                num nSigType[3]
                num nValue[3]
            mdesc mMdesc = {leave=0}
            num nActionIndex = 60
            num nDelay = 1
            num nMoveType = 1
            num nPercentage
            num nSigValue = 1
        pointRx pPointRx[2] = {x=-138.850367, y=-44.569058, z=962.511805, rx=-1.752214, ry=-0.122124, rz=-89.326646, shoulder=lefty, elbow=epositive, wrist=wpositive}
        string sID
      [75]
        bool bMarked
        jointRx jJointRx = {j1=-49.904251, j2=-65.605747, j3=139.0621971, j4=-181.0710428, j5=74.878861, j6=140.871685}
        pointRx pInter
        paraItem pParaItem
          [0]
            bool bSafePoint
            ifItem iIfItem
              [0]
                bool bANDOR[2]
                num nSigIndex[3]
                num nSigType[3]
                num nValue[3]
            mdesc mMdesc = {leave=0}
            num nActionIndex = 60
            num nDelay = 1
            num nMoveType = 1
            num nPercentage
            num nSigValue = 1
        pointRx pPointRx[2] = {x=-44.539892, y=-44.568217, z=962.547058, rx=-1.752061, ry=-0.123361, rz=-89.326689, shoulder=lefty, elbow=epositive, wrist=wpositive}
        string sID
      [76]
        bool bMarked
        jointRx jJointRx = {j1=-49.289261, j2=-63.229169, j3=134.202102, j4=-181.102758, j5=72.384398, j6=140.311025}
        pointRx pInter
        paraItem pParaItem
          [0]
            bool bSafePoint
            ifItem iIfItem
              [0]
                bool bANDOR[2]
                num nSigIndex[3]
                num nSigType[3]
                num nValue[3]
            mdesc mMdesc = {leave=0}
            num nActionIndex = 60
            num nDelay = 1
            num nMoveType = 1
            num nPercentage
            num nSigValue = 1
        pointRx pPointRx[2] = {x=-42.782853, y=-44.569273, z=1003.955298, rx=-1.753071, ry=-0.121713, rz=-89.326781, shoulder=lefty, elbow=epositive, wrist=wpositive}
        string sID
      [77]
        bool bMarked
        jointRx jJointRx = {j1=-25.432487, j2=-45.494499, j3=127.259364, j4=-181.493414, j5=82.715062, j6=116.303511}
        pointRx pInter
        paraItem pParaItem
          [0]
            bool bSafePoint
            ifItem iIfItem
              [0]
                bool bANDOR[2]
                num nSigIndex[3]
                num nSigType[3]
                num nValue[3]
            mdesc mMdesc = {leave=0}
            num nActionIndex = 60
            num nDelay = 1
            num nMoveType = 1
            num nPercentage
            num nSigValue = 1
        pointRx pPointRx[2] = {x=73.884399, y=-40.550183, z=1028.430042, rx=-1.744787, ry=-0.219486, rz=-89.333983, shoulder=lefty, elbow=epositive, wrist=wpositive}
        string sID
      [78]
        bool bMarked
        jointRx jJointRx = {j1=-57.856377, j2=-66.18455, j3=133.138862, j4=-180.798841, j5=68.549304, j6=148.828951}
        pointRx pInter
        paraItem pParaItem
          [0]
            bool bSafePoint
            ifItem iIfItem
              [0]
                bool bANDOR[2]
                num nSigIndex[3]
                num nSigType[3]
                num nValue[3]
            mdesc mMdesc = {leave=0}
            num nActionIndex = 60
            num nDelay = 1
            num nMoveType = 1
            num nPercentage
            num nSigValue = 1
        pointRx pPointRx[2] = {x=-67.43152, y=-40.567065, z=1016.367875, rx=-1.744462, ry=-0.217896, rz=-89.333233, shoulder=lefty, elbow=epositive, wrist=wpositive}
        string sID
      [79]
        bool bMarked
        jointRx jJointRx = {j1=-125.666138, j2=-76.447258, j3=135.218346, j4=-178.621352, j5=60.0693288, j6=215.6343}
        pointRx pInter
        paraItem pParaItem
          [0]
            bool bSafePoint
            ifItem iIfItem
              [0]
                bool bANDOR[2]
                num nSigIndex[3]
                num nSigType[3]
                num nValue[3]
            mdesc mMdesc = {leave=0}
            num nActionIndex = 60
            num nDelay = 1
            num nMoveType = 1
            num nPercentage
            num nSigValue = 1
        pointRx pPointRx[2] = {x=-141.607559, y=-40.56496, z=1001.487797, rx=-1.745427, ry=-0.218033, rz=-89.333718, shoulder=lefty, elbow=epositive, wrist=wpositive}
        string sID
      [80]
        bool bMarked
        jointRx jJointRx = {j1=-163.468753, j2=-72.941717, j3=129.657925, j4=-177.930129, j5=57.0209808, j6=253.00669774}
        pointRx pInter
        paraItem pParaItem
          [0]
            bool bSafePoint
            ifItem iIfItem
              [0]
                bool bANDOR[2]
                num nSigIndex[3]
                num nSigType[3]
                num nValue[3]
            mdesc mMdesc = {leave=0}
            num nActionIndex = 60
            num nDelay = 1
            num nMoveType = 1
            num nPercentage
            num nSigValue = 1
        pointRx pPointRx[2] = {x=-178.509464, y=-40.567787, z=1047.669101, rx=-1.746323, ry=-0.218277, rz=-89.333981, shoulder=lefty, elbow=epositive, wrist=wpositive}
        string sID
      [81]
        bool bMarked
        jointRx jJointRx = {j1=-177.244487, j2=-58.712757, j3=130.795458, j4=-178.155232, j5=71.95685, j6=267.344536}
        pointRx pInter
        paraItem pParaItem
          [0]
            bool bSafePoint
            ifItem iIfItem
              [0]
                bool bANDOR[2]
                num nSigIndex[3]
                num nSigType[3]
                num nValue[3]
            mdesc mMdesc = {leave=0}
            num nActionIndex = 60
            num nDelay = 1
            num nMoveType = 1
            num nPercentage
            num nSigValue = 1
        pointRx pPointRx[2] = {x=-305.74421, y=-40.564807, z=1028.0320815, rx=-1.745533, ry=-0.218693, rz=-89.333779, shoulder=lefty, elbow=epositive, wrist=wpositive}
        string sID
      [82]
        bool bMarked
        jointRx jJointRx = {j1=-178.526843, j2=-40.454962, j3=125.405301, j4=-178.242312, j5=84.778901, j6=269.0391142}
        pointRx pInter
        paraItem pParaItem
          [0]
            bool bSafePoint
            ifItem iIfItem
              [0]
                bool bANDOR[2]
                num nSigIndex[3]
                num nSigType[3]
                num nValue[3]
            mdesc mMdesc = {leave=0}
            num nActionIndex = 60
            num nDelay = 1
            num nMoveType = 1
            num nPercentage
            num nSigValue = 1
        pointRx pPointRx[2] = {x=-434.343088, y=-40.61718, z=1028.0320848, rx=-1.745356, ry=-0.218738, rz=-89.333719, shoulder=lefty, elbow=epositive, wrist=wpositive}
        string sID
      [83]
        bool bMarked
        jointRx jJointRx = {j1=-178.966416, j2=-24.85944, j3=117.444048, j4=-178.24946, j5=92.396091, j6=269.712104}
        pointRx pInter
        paraItem pParaItem
          [0]
            bool bSafePoint
            ifItem iIfItem
              [0]
                bool bANDOR[2]
                num nSigIndex[3]
                num nSigType[3]
                num nValue[3]
            mdesc mMdesc = {leave=0}
            num nActionIndex = 60
            num nDelay = 1
            num nMoveType = 1
            num nPercentage
            num nSigValue = 1
        pointRx pPointRx[2] = {x=-550.558, y=-40.617172, z=1028.0320539, rx=-1.745357, ry=-0.218827, rz=-89.333714, shoulder=lefty, elbow=epositive, wrist=wpositive}
        string sID
      [84]
        bool bMarked
        jointRx jJointRx = {j1=-178.990337, j2=-23.604156, j3=109.459463, j4=-178.246238, j5=85.670511, j6=269.530325}
        pointRx pInter
        paraItem pParaItem
          [0]
            bool bSafePoint
            ifItem iIfItem
              [0]
                bool bANDOR[2]
                num nSigIndex[3]
                num nSigType[3]
                num nValue[3]
            mdesc mMdesc = {leave=0}
            num nActionIndex = 60
            num nDelay = 1
            num nMoveType = 1
            num nPercentage
            num nSigValue = 1
        pointRx pPointRx[2] = {x=-559.676751, y=-40.616999, z=1097.0852879, rx=-1.745205, ry=-0.217512, rz=-89.33374, shoulder=lefty, elbow=epositive, wrist=wpositive}
        string sID
      [85]
        bool bMarked
        jointRx jJointRx = {j1=-178.943744, j2=-24.322013, j3=101.711175, j4=-178.206641, j5=77.210582, j6=269.219034}
        pointRx pInter
        paraItem pParaItem
          [0]
            bool bSafePoint
            ifItem iIfItem
              [0]
                bool bANDOR[2]
                num nSigIndex[3]
                num nSigType[3]
                num nValue[3]
            mdesc mMdesc = {leave=0}
            num nActionIndex = 60
            num nDelay = 1
            num nMoveType = 1
            num nPercentage
            num nSigValue = 1
        pointRx pPointRx[2] = {x=-542.070783, y=-40.616994, z=1174.87195, rx=-1.745164, ry=-0.216758, rz=-89.333713, shoulder=lefty, elbow=epositive, wrist=wpositive}
        string sID
      [86]
        bool bMarked
        jointRx jJointRx = {j1=-178.943806, j2=-23.793943, j3=99.30263, j4=-178.192287, j5=75.331347, j6=269.158327}
        pointRx pInter
        paraItem pParaItem
          [0]
            bool bSafePoint
            ifItem iIfItem
              [0]
                bool bANDOR[2]
                num nSigIndex[3]
                num nSigType[3]
                num nValue[3]
            mdesc mMdesc = {leave=0}
            num nActionIndex = 60
            num nDelay = 1
            num nMoveType = 1
            num nPercentage
            num nSigValue = 1
        pointRx pPointRx[2] = {x=-542.046055, y=-40.616997, z=1194.299438, rx=-1.745092, ry=-0.216442, rz=-89.333682, shoulder=lefty, elbow=epositive, wrist=wpositive}
        string sID
      [87]
        bool bMarked
        jointRx jJointRx = {j1=-178.85922, j2=-27.330123, j3=102.744036, j4=-178.191054, j5=75.238753, j6=269.0705123}
        pointRx pInter
        paraItem pParaItem
          [0]
            bool bSafePoint
            ifItem iIfItem
              [0]
                bool bANDOR[2]
                num nSigIndex[3]
                num nSigType[3]
                num nValue[3]
            mdesc mMdesc = {leave=0}
            num nActionIndex = 60
            num nDelay = 1
            num nMoveType = 1
            num nPercentage
            num nSigValue = 1
        pointRx pPointRx[2] = {x=-513.909364, y=-40.617001, z=1181.865557, rx=-1.745263, ry=-0.216897, rz=-89.333745, shoulder=lefty, elbow=epositive, wrist=wpositive}
        string sID
      [88]
        bool bMarked
        jointRx jJointRx = {j1=-178.577868, j2=-35.0352996, j3=106.0927297, j4=-178.147828, j5=70.89347, j6=268.643627}
        pointRx pInter
        paraItem pParaItem
          [0]
            bool bSafePoint
            ifItem iIfItem
              [0]
                bool bANDOR[2]
                num nSigIndex[3]
                num nSigType[3]
                num nValue[3]
            mdesc mMdesc = {leave=0}
            num nActionIndex = 60
            num nDelay = 1
            num nMoveType = 1
            num nPercentage
            num nSigValue = 1
        pointRx pPointRx[2] = {x=-444.101189, y=-40.617001, z=1187.110134, rx=-1.745281, ry=-0.216517, rz=-89.333733, shoulder=lefty, elbow=epositive, wrist=wpositive}
        string sID
      [89]
        bool bMarked
        jointRx jJointRx = {j1=-177.964362, j2=-47.427804, j3=117.345153, j4=-178.132839, j5=69.773165, j6=267.990525}
        pointRx pInter
        paraItem pParaItem
          [0]
            bool bSafePoint
            ifItem iIfItem
              [0]
                bool bANDOR[2]
                num nSigIndex[3]
                num nSigType[3]
                num nValue[3]
            mdesc mMdesc = {leave=0}
            num nActionIndex = 60
            num nDelay = 1
            num nMoveType = 1
            num nPercentage
            num nSigValue = 1
        pointRx pPointRx[2] = {x=-358.696243, y=-40.617001, z=1126.286618, rx=-1.745413, ry=-0.216112, rz=-89.333736, shoulder=lefty, elbow=epositive, wrist=wpositive}
        string sID
      [90]
        bool bMarked
        jointRx jJointRx = {j1=-177.960401, j2=-42.42338, j3=104.324192, j4=-178.0116171, j5=61.761954, j6=267.691309}
        pointRx pInter
        paraItem pParaItem
          [0]
            bool bSafePoint
            ifItem iIfItem
              [0]
                bool bANDOR[2]
                num nSigIndex[3]
                num nSigType[3]
                num nValue[3]
            mdesc mMdesc = {leave=0}
            num nActionIndex = 60
            num nDelay = 1
            num nMoveType = 1
            num nPercentage
            num nSigValue = 1
        pointRx pPointRx[2] = {x=-358.210554, y=-40.616999, z=1227.312647, rx=-1.745114, ry=-0.215409, rz=-89.333647, shoulder=lefty, elbow=epositive, wrist=wpositive}
        string sID
      [91]
        bool bMarked
        jointRx jJointRx = {j1=-157.648785, j2=-55.0873266, j3=110.653004, j4=-177.95404, j5=56.0449416, j6=247.169842}
        pointRx pInter
        paraItem pParaItem
          [0]
            bool bSafePoint
            ifItem iIfItem
              [0]
                bool bANDOR[2]
                num nSigIndex[3]
                num nSigType[3]
                num nValue[3]
            mdesc mMdesc = {leave=0}
            num nActionIndex = 60
            num nDelay = 1
            num nMoveType = 1
            num nPercentage
            num nSigValue = 1
        pointRx pPointRx[2] = {x=-229.83526, y=-65.451897, z=1196.333444, rx=-1.745262, ry=-0.217825, rz=-89.332323, shoulder=lefty, elbow=epositive, wrist=wpositive}
        string sID
      [92]
        bool bMarked
        jointRx jJointRx = {j1=-152.966394, j2=-56.240625, j3=110.746536, j4=-177.982817, j5=55.121987, j6=242.474574}
        pointRx pInter
        paraItem pParaItem
          [0]
            bool bSafePoint
            ifItem iIfItem
              [0]
                bool bANDOR[2]
                num nSigIndex[3]
                num nSigType[3]
                num nValue[3]
            mdesc mMdesc = {leave=0}
            num nActionIndex = 60
            num nDelay = 1
            num nMoveType = 1
            num nPercentage
            num nSigValue = 1
        pointRx pPointRx[2] = {x=-212.6845, y=-65.452346, z=1196.358042, rx=-1.746333, ry=-0.218302, rz=-89.332682, shoulder=lefty, elbow=epositive, wrist=wpositive}
        string sID
      [93]
        bool bMarked
        jointRx jJointRx = {j1=-118.542599, j2=-58.519116, j3=112.0638486, j4=-178.749072, j5=54.980609, j6=208.482941}
        pointRx pInter
        paraItem pParaItem
          [0]
            bool bSafePoint
            ifItem iIfItem
              [0]
                bool bANDOR[2]
                num nSigIndex[3]
                num nSigType[3]
                num nValue[3]
            mdesc mMdesc = {leave=0}
            num nActionIndex = 60
            num nDelay = 1
            num nMoveType = 1
            num nPercentage
            num nSigValue = 1
        pointRx pPointRx[2] = {x=-149.858699, y=-65.452346, z=1187.0826994, rx=-1.745135, ry=-0.217044, rz=-89.332258, shoulder=lefty, elbow=epositive, wrist=wpositive}
        string sID
      [94]
        bool bMarked
        jointRx jJointRx = {j1=-101.200662, j2=-58.679642, j3=113.706302, j4=-179.339305, j5=56.697308, j6=191.500759}
        pointRx pInter
        paraItem pParaItem
          [0]
            bool bSafePoint
            ifItem iIfItem
              [0]
                bool bANDOR[2]
                num nSigIndex[3]
                num nSigType[3]
                num nValue[3]
            mdesc mMdesc = {leave=0}
            num nActionIndex = 60
            num nDelay = 1
            num nMoveType = 1
            num nPercentage
            num nSigValue = 1
        pointRx pPointRx[2] = {x=-127.503998, y=-65.472867, z=1174.335896, rx=-1.744346, ry=-0.217552, rz=-89.332398, shoulder=lefty, elbow=epositive, wrist=wpositive}
        string sID
      [95]
        bool bMarked
        jointRx jJointRx = {j1=-101.203749, j2=-57.0328969, j3=110.693044, j4=-179.328951, j5=55.331019, j6=191.484931}
        pointRx pInter
        paraItem pParaItem
          [0]
            bool bSafePoint
            ifItem iIfItem
              [0]
                bool bANDOR[2]
                num nSigIndex[3]
                num nSigType[3]
                num nValue[3]
            mdesc mMdesc = {leave=0}
            num nActionIndex = 60
            num nDelay = 1
            num nMoveType = 1
            num nPercentage
            num nSigValue = 1
        pointRx pPointRx[2] = {x=-127.503988, y=-65.473043, z=1197.162512, rx=-1.744433, ry=-0.217146, rz=-89.332357, shoulder=lefty, elbow=epositive, wrist=wpositive}
        string sID
      [96]
        bool bMarked
        jointRx jJointRx = {j1=-84.916197, j2=-57.654127, j3=112.0354709, j4=-179.926433, j5=56.138092, j6=175.545215}
        pointRx pInter
        paraItem pParaItem
          [0]
            bool bSafePoint
            ifItem iIfItem
              [0]
                bool bANDOR[2]
                num nSigIndex[3]
                num nSigType[3]
                num nValue[3]
            mdesc mMdesc = {leave=0}
            num nActionIndex = 60
            num nDelay = 1
            num nMoveType = 1
            num nPercentage
            num nSigValue = 1
        pointRx pPointRx[2] = {x=-105.833813, y=-53.577317, z=1186.997866, rx=-1.744409, ry=-0.216493, rz=-89.33235, shoulder=lefty, elbow=epositive, wrist=wpositive}
        string sID
      [97]
        bool bMarked
        jointRx jJointRx = {j1=-74.942351, j2=-49.0636516, j3=113.425459, j4=-183.373141, j5=77.590842, j6=166.743204}
        pointRx pInter
        paraItem pParaItem
          [0]
            bool bSafePoint
            ifItem iIfItem
              [0]
                bool bANDOR[2]
                num nSigIndex[3]
                num nSigType[3]
                num nValue[3]
            mdesc mMdesc = {leave=0}
            num nActionIndex = 60
            num nDelay = 1
            num nMoveType = 1
            num nPercentage
            num nSigValue = 1
        pointRx pPointRx[2] = {x=-70.288394, y=-10.197743, z=1148.602795, rx=-13.604008, ry=-0.216042, rz=-89.332075, shoulder=lefty, elbow=epositive, wrist=wpositive}
        string sID
      [98]
        bool bMarked
        jointRx jJointRx = {j1=-22.441628, j2=-49.998667, j3=113.146837, j4=-179.268601, j5=63.114949, j6=112.777772}
        pointRx pInter
        paraItem pParaItem
          [0]
            bool bSafePoint
            ifItem iIfItem
              [0]
                bool bANDOR[2]
                num nSigIndex[3]
                num nSigType[3]
                num nValue[3]
            mdesc mMdesc = {leave=0}
            num nActionIndex = 60
            num nDelay = 1
            num nMoveType = 1
            num nPercentage
            num nSigValue = 1
        pointRx pPointRx[2] = {x=2.572536, y=-22.293277, z=1169.165569, rx=0.616343, ry=-0.216579, rz=-89.332136, shoulder=lefty, elbow=epositive, wrist=wpositive}
        string sID
      [99]
        bool bMarked
        jointRx jJointRx = {j1=-16.222078, j2=-42.747965, j3=111.131068, j4=-179.299489, j5=68.420107, j6=106.63085}
        pointRx pInter
        paraItem pParaItem
          [0]
            bool bSafePoint
            ifItem iIfItem
              [0]
                bool bANDOR[2]
                num nSigIndex[3]
                num nSigType[3]
                num nValue[3]
            mdesc mMdesc = {leave=0}
            num nActionIndex = 60
            num nDelay = 1
            num nMoveType = 1
            num nPercentage
            num nSigValue = 1
        pointRx pPointRx[2] = {x=64.811204, y=-22.293322, z=1169.130311, rx=0.615547, ry=-0.216097, rz=-89.332208, shoulder=lefty, elbow=epositive, wrist=wpositive}
        string sID
      [100]
        bool bMarked
        jointRx jJointRx = {j1=-11.927651, j2=-32.0900118, j3=103.0810682, j4=-179.315894, j5=71.0760377, j6=102.371735}
        pointRx pInter
        paraItem pParaItem
          [0]
            bool bSafePoint
            ifItem iIfItem
              [0]
                bool bANDOR[2]
                num nSigIndex[3]
                num nSigType[3]
                num nValue[3]
            mdesc mMdesc = {leave=0}
            num nActionIndex = 60
            num nDelay = 1
            num nMoveType = 1
            num nPercentage
            num nSigValue = 1
        pointRx pPointRx[2] = {x=145.897455, y=-22.29476, z=1202.0898265, rx=0.615855, ry=-0.215659, rz=-89.332409, shoulder=lefty, elbow=epositive, wrist=wpositive}
        string sID
      [101]
        bool bMarked
        jointRx jJointRx = {j1=-14.974019, j2=-36.733975, j3=99.744873, j4=-179.269184, j5=63.0625851, j6=105.309151}
        pointRx pInter
        paraItem pParaItem
          [0]
            bool bSafePoint
            ifItem iIfItem
              [0]
                bool bANDOR[2]
                num nSigIndex[3]
                num nSigType[3]
                num nValue[3]
            mdesc mMdesc = {leave=0}
            num nActionIndex = 60
            num nDelay = 1
            num nMoveType = 1
            num nPercentage
            num nSigValue = 1
        pointRx pPointRx[2] = {x=83.529929, y=-22.294757, z=1249.648683, rx=0.616531, ry=-0.216447, rz=-89.332334, shoulder=lefty, elbow=epositive, wrist=wpositive}
        string sID
      [102]
        bool bMarked
        jointRx jJointRx = {j1=-14.974848, j2=-34.297369, j3=93.572735, j4=-179.243247, j5=59.326428, j6=105.254901}
        pointRx pInter
        paraItem pParaItem
          [0]
            bool bSafePoint
            ifItem iIfItem
              [0]
                bool bANDOR[2]
                num nSigIndex[3]
                num nSigType[3]
                num nValue[3]
            mdesc mMdesc = {leave=0}
            num nActionIndex = 60
            num nDelay = 1
            num nMoveType = 1
            num nPercentage
            num nSigValue = 1
        pointRx pPointRx[2] = {x=83.543818, y=-22.294762, z=1293.403623, rx=0.616141, ry=-0.215384, rz=-89.33244, shoulder=lefty, elbow=epositive, wrist=wpositive}
        string sID
      [103]
        bool bMarked
        jointRx jJointRx = {j1=-45.0792437, j2=-47.932825, j3=93.769334, j4=-179.178005, j5=45.55525, j6=135.171407}
        pointRx pInter
        paraItem pParaItem
          [0]
            bool bSafePoint
            ifItem iIfItem
              [0]
                bool bANDOR[2]
                num nSigIndex[3]
                num nSigType[3]
                num nValue[3]
            mdesc mMdesc = {leave=0}
            num nActionIndex = 60
            num nDelay = 1
            num nMoveType = 1
            num nPercentage
            num nSigValue = 1
        pointRx pPointRx[2] = {x=-75.0284555, y=-24.9462, z=1317.531429, rx=0.61562, ry=-0.214846, rz=-89.332539, shoulder=lefty, elbow=epositive, wrist=wpositive}
        string sID
      [104]
        bool bMarked
        jointRx jJointRx = {j1=-104.199394, j2=-58.872088, j3=119.262884, j4=-178.287616, j5=65.702617, j6=194.100128}
        pointRx pInter
        paraItem pParaItem
          [0]
            bool bSafePoint
            ifItem iIfItem
              [0]
                bool bANDOR[2]
                num nSigIndex[3]
                num nSigType[3]
                num nValue[3]
            mdesc mMdesc = {leave=0}
            num nActionIndex = 60
            num nDelay = 1
            num nMoveType = 1
            num nPercentage
            num nSigValue = 1
        pointRx pPointRx[2] = {x=-138.333641, y=-53.548008, z=1127.0142429, rx=-5.522356, ry=-0.214514, rz=-89.33257, shoulder=lefty, elbow=epositive, wrist=wpositive}
        string sID
      [105]
        bool bMarked
        jointRx jJointRx = {j1=-168.930499, j2=-33.269754, j3=111.495151, j4=-174.438533, j5=79.127174, j6=258.515266}
        pointRx pInter
        paraItem pParaItem
          [0]
            bool bSafePoint
            ifItem iIfItem
              [0]
                bool bANDOR[2]
                num nSigIndex[3]
                num nSigType[3]
                num nValue[3]
            mdesc mMdesc = {leave=0}
            num nActionIndex = 60
            num nDelay = 1
            num nMoveType = 1
            num nPercentage
            num nSigValue = 1
        pointRx pPointRx[2] = {x=-460.931799, y=-53.549955, z=1127.0747297, rx=-5.522947, ry=-0.215065, rz=-89.332743, shoulder=lefty, elbow=epositive, wrist=wpositive}
        string sID
      [106]
        bool bMarked
        jointRx jJointRx = {j1=-178.718432, j2=-47.656061, j3=94.0601296, j4=-179.783558, j5=46.19183, j6=269.235916}
        pointRx pInter
        paraItem pParaItem
          [0]
            bool bSafePoint
            ifItem iIfItem
              [0]
                bool bANDOR[2]
                num nSigIndex[3]
                num nSigType[3]
                num nValue[3]
            mdesc mMdesc = {leave=0}
            num nActionIndex = 60
            num nDelay = 1
            num nMoveType = 1
            num nPercentage
            num nSigValue = 1
        pointRx pPointRx[2] = {x=-239.874829, y=-52.0270152, z=1315.44798, rx=-0.151408, ry=-0.215882, rz=-89.333259, shoulder=lefty, elbow=epositive, wrist=wpositive}
        string sID
      [107]
        bool bMarked
        jointRx jJointRx = {j1=-174.208935, j2=-36.617887, j3=92.316666, j4=-177.741125, j5=55.691456, j6=263.60606}
        pointRx pInter
        paraItem pParaItem
          [0]
            bool bSafePoint
            ifItem iIfItem
              [0]
                bool bANDOR[2]
                num nSigIndex[3]
                num nSigType[3]
                num nValue[3]
            mdesc mMdesc = {leave=0}
            num nActionIndex = 60
            num nDelay = 1
            num nMoveType = 1
            num nPercentage
            num nSigValue = 1
        pointRx pPointRx[2] = {x=-362.264063, y=-53.0173082, z=1310.403557, rx=-1.853366, ry=-0.216126, rz=-89.333164, shoulder=lefty, elbow=epositive, wrist=wpositive}
        string sID
      [108]
        bool bMarked
        jointRx jJointRx = {j1=-174.64878, j2=-31.90972, j3=92.577201, j4=-177.85981, j5=60.641464, j6=264.270204}
        pointRx pInter
        paraItem pParaItem
          [0]
            bool bSafePoint
            ifItem iIfItem
              [0]
                bool bANDOR[2]
                num nSigIndex[3]
                num nSigType[3]
                num nValue[3]
            mdesc mMdesc = {leave=0}
            num nActionIndex = 60
            num nDelay = 1
            num nMoveType = 1
            num nPercentage
            num nSigValue = 1
        pointRx pPointRx[2] = {x=-421.633734, y=-56.993181, z=1293.0105914, rx=-1.85308, ry=-0.216814, rz=-89.333136, shoulder=lefty, elbow=epositive, wrist=wpositive}
        string sID
      [109]
        bool bMarked
        jointRx jJointRx = {j1=-176.308868, j2=-19.882778, j3=85.885827, j4=-177.959065, j5=65.918849, j6=266.147536}
        pointRx pInter
        paraItem pParaItem
          [0]
            bool bSafePoint
            ifItem iIfItem
              [0]
                bool bANDOR[2]
                num nSigIndex[3]
                num nSigType[3]
                num nValue[3]
            mdesc mMdesc = {leave=0}
            num nActionIndex = 60
            num nDelay = 1
            num nMoveType = 1
            num nPercentage
            num nSigValue = 1
        pointRx pPointRx[2] = {x=-540.666158, y=-56.993339, z=1293.00889756, rx=-1.853097, ry=-0.217424, rz=-89.333381, shoulder=lefty, elbow=epositive, wrist=wpositive}
        string sID
      [110]
        bool bMarked
        jointRx jJointRx = {j1=-176.149742, j2=-21.522794, j3=86.947142, j4=-177.949917, j5=65.34723, j6=265.966515}
        pointRx pInter
        paraItem pParaItem
          [0]
            bool bSafePoint
            ifItem iIfItem
              [0]
                bool bANDOR[2]
                num nSigIndex[3]
                num nSigType[3]
                num nValue[3]
            mdesc mMdesc = {leave=0}
            num nActionIndex = 60
            num nDelay = 1
            num nMoveType = 1
            num nPercentage
            num nSigValue = 1
        pointRx pPointRx[2] = {x=-524.804732, y=-56.995789, z=1293.0175935, rx=-1.852848, ry=-0.215861, rz=-89.332769, shoulder=lefty, elbow=epositive, wrist=wpositive}
        string sID
      [111]
        bool bMarked
        jointRx jJointRx = {j1=-176.379023, j2=-14.996563, j3=73.511352, j4=-177.814157, j5=58.436024, j6=265.907384}
        pointRx pInter
        paraItem pParaItem
          [0]
            bool bSafePoint
            ifItem iIfItem
              [0]
                bool bANDOR[2]
                num nSigIndex[3]
                num nSigType[3]
                num nValue[3]
            mdesc mMdesc = {leave=0}
            num nActionIndex = 60
            num nDelay = 1
            num nMoveType = 1
            num nPercentage
            num nSigValue = 1
        pointRx pPointRx[2] = {x=-547.946589, y=-56.996452, z=1369.367078, rx=-1.852482, ry=-0.21472, rz=-89.33211, shoulder=lefty, elbow=epositive, wrist=wpositive}
        string sID
      [112]
        bool bMarked
        jointRx jJointRx = {j1=-174.680222, j2=-27.0244183, j3=80.825627, j4=-177.689262, j5=53.783296, j6=263.986809}
        pointRx pInter
        paraItem pParaItem
          [0]
            bool bSafePoint
            ifItem iIfItem
              [0]
                bool bANDOR[2]
                num nSigIndex[3]
                num nSigType[3]
                num nValue[3]
            mdesc mMdesc = {leave=0}
            num nActionIndex = 60
            num nDelay = 1
            num nMoveType = 1
            num nPercentage
            num nSigValue = 1
        pointRx pPointRx[2] = {x=-423.0814867, y=-56.996861, z=1369.379158, rx=-1.852359, ry=-0.212738, rz=-89.331744, shoulder=lefty, elbow=epositive, wrist=wpositive}
        string sID
      [113]
        bool bMarked
        jointRx jJointRx = {j1=-174.323366, j2=-28.55257, j3=81.546918, j4=-177.665438, j5=52.989259, j6=263.590154}
        pointRx pInter
        paraItem pParaItem
          [0]
            bool bSafePoint
            ifItem iIfItem
              [0]
                bool bANDOR[2]
                num nSigIndex[3]
                num nSigType[3]
                num nValue[3]
            mdesc mMdesc = {leave=0}
            num nActionIndex = 60
            num nDelay = 1
            num nMoveType
            num nPercentage
            num nSigValue = 1
        pointRx pPointRx[2] = {x=-406.271248, y=-57.000225416, z=1369.381759, rx=-1.852116, ry=-0.212153, rz=-89.331276, shoulder=lefty, elbow=epositive, wrist=wpositive}
        string sID
      [114]
        bool bMarked
        jointRx jJointRx = {j1=-175.249593, j2=-37.427588, j3=140.969865, j4=-180.67062, j5=122.873549, j6=265.286535}
        pointRx pInter
        paraItem pParaItem
          [0]
            bool bSafePoint
            ifItem iIfItem
              [0]
                bool bANDOR[2]
                num nSigIndex[3]
                num nSigType[3]
                num nValue[3]
            mdesc mMdesc = {leave=0}
            num nActionIndex = 60
            num nDelay = 1
            num nMoveType
            num nPercentage
            num nSigValue = 1
        pointRx pPointRx[2] = {x=-228.283263, y=-62.885699, z=887.339634, rx=-1.0697557, ry=19.312473, rz=-89.512958, shoulder=lefty, elbow=epositive, wrist=wpositive}
        string sID
      [115]
        bool bMarked
        jointRx jJointRx = {j1=-55.114066, j2=-37.427631, j3=140.969917, j4=-194.186695, j5=122.873144, j6=139.0711954}
        pointRx pInter
        paraItem pParaItem
          [0]
            bool bSafePoint
            ifItem iIfItem
              [0]
                bool bANDOR[2]
                num nSigIndex[3]
                num nSigType[3]
                num nValue[3]
            mdesc mMdesc = {leave=0}
            num nActionIndex = 60
            num nDelay = 1
            num nMoveType
            num nPercentage
            num nSigValue = 1
        pointRx pPointRx[2] = {x=27.342979, y=34.851056, z=815.295742, rx=-23.222086, ry=-1.370042, rz=-90.628941, shoulder=lefty, elbow=epositive, wrist=wpositive}
        string sID
      [116]
        bool bMarked
        jointRx jJointRx = {j1=13.421796, j2=-4.818794, j3=127.476333, j4=-178.119312, j5=122.0945871, j6=-9.799703}
        pointRx pInter
        paraItem pParaItem
          [0]
            bool bSafePoint
            ifItem iIfItem
              [0]
                bool bANDOR[2]
                num nSigIndex[3]
                num nSigType[3]
                num nValue[3]
            mdesc mMdesc = {leave=0}
            num nActionIndex = 60
            num nDelay = 1
            num nMoveType = 1
            num nPercentage
            num nSigValue = 1
        pointRx pPointRx[2] = {x=448.772207, y=302.863979, z=805.266279, rx=1.422401, ry=0.903641, rz=-177.39626, shoulder=lefty, elbow=epositive, wrist=wpositive}
        string sID
      [117]
        bool bMarked
        jointRx jJointRx = {j1=-0.745998, j2=38.655383, j3=103.0614514, j4=-179.633274, j5=123.453989, j6=8.386247}
        pointRx pInter
        paraItem pParaItem
          [0]
            bool bSafePoint
            ifItem iIfItem
              [0]
                bool bANDOR[2]
                num nSigIndex[3]
                num nSigType[3]
                num nValue[3]
            mdesc mMdesc = {leave=0}
            num nActionIndex = 60
            num nDelay = 1
            num nMoveType = 1
            num nPercentage
            num nSigValue = 1
        pointRx pPointRx[2] = {x=872.320063, y=193.823231, z=536.442949, rx=0.568319, ry=18.256239, rz=-172.702412, shoulder=lefty, elbow=epositive, wrist=wpositive}
        string sID
    string sID
  [PRO2-BlowPATH]
    num nFrameIndex
    num nMoveID
    num nToolIndex
    pointItem pPointItem
      [0]
        bool bMarked
        jointRx jJointRx = {j1=25.205089, j2=131.889625, j3=-138.179149, j4=-50.606575, j5=-24.632261, j6=111.315059}
        pointRx pInter
        paraItem pParaItem
          [0]
            bool bSafePoint
            ifItem iIfItem
              [0]
                bool bANDOR[2]
                num nSigIndex[3]
                num nSigType[3]
                num nValue[3]
            mdesc mMdesc
            num nActionIndex = 60
            num nDelay = 1
            num nMoveType = 7
            num nPercentage
            num nSigValue = 1
        pointRx pPointRx[2] = {x=93.0356449, y=143.591414, z=599.882332, rx=84.531042, ry=-6.510159, rz=117.916178, shoulder=lefty, elbow=enegative, wrist=wnegative}
        string sID
    string sID
  [Position5_point_blow]
    num nFrameIndex
    num nMoveID
    num nToolIndex
    pointItem pPointItem[48]
      [0]
        bool bMarked
        jointRx jJointRx
        pointRx pInter
        paraItem pParaItem
          [0]
            bool bSafePoint
            ifItem iIfItem
              [0]
                bool bANDOR[2]
                num nSigIndex[3]
                num nSigType[3]
                num nValue[3]
            mdesc mMdesc
            num nActionIndex = 43
            num nDelay
            num nMoveType = 4
            num nPercentage
            num nSigValue = 1
        pointRx pPointRx[2]
        string sID
      [1]
        bool bMarked
        jointRx jJointRx = {j1=-87.551314, j2=145.129335, j3=-83.0857287, j4=182.11845, j5=63.691242, j6=-64.966659}
        pointRx pInter
        paraItem pParaItem
          [0]
            bool bSafePoint
            ifItem iIfItem
              [0]
                bool bANDOR[2]
                num nSigIndex[3]
                num nSigType[3]
                num nValue[3]
            mdesc mMdesc
            num nActionIndex = 42
            num nDelay
            num nMoveType = 1
            num nPercentage
            num nSigValue = 1
        pointRx pPointRx[2] = {x=61.349727, y=-652.129552, z=350.0734551, rx=-1.549449, ry=-1.96692, rz=28.421736, shoulder=lefty, elbow=enegative, wrist=wpositive}
        string sID
      [2]
        bool bMarked
        jointRx jJointRx = {j1=-47.00566362, j2=123.661152, j3=-79.978164, j4=176.739672, j5=50.379836, j6=-102.275032}
        pointRx pInter
        paraItem pParaItem
          [0]
            bool bSafePoint
            ifItem iIfItem
              [0]
                bool bANDOR[2]
                num nSigIndex[3]
                num nSigType[3]
                num nValue[3]
            mdesc mMdesc
            num nActionIndex = 42
            num nDelay
            num nMoveType = 1
            num nPercentage
            num nSigValue = 1
        pointRx pPointRx[2] = {x=488.627273, y=-418.649607, z=567.937104, rx=-6.582637, ry=-2.686226, rz=28.338446, shoulder=lefty, elbow=enegative, wrist=wpositive}
        string sID
      [3]
        bool bMarked
        jointRx jJointRx = {j1=-49.0942088, j2=121.00459063, j3=-74.169176, j4=177.183335, j5=53.609232, j6=-100.608132}
        pointRx pInter
        paraItem pParaItem
          [0]
            bool bSafePoint
            ifItem iIfItem
              [0]
                bool bANDOR[2]
                num nSigIndex[3]
                num nSigType[3]
                num nValue[3]
            mdesc mMdesc
            num nActionIndex = 42
            num nDelay
            num nMoveType = 1
